ABB RAPID module: CalibData.mod

MODULE CalibData
    PERS tooldata My_Mechanism_1:=[TRUE,[[0,0,90],[1,0,0,0]],[1,[0,0,90],[1,0,0,0],0,0,0]];
    TASK PERS wobjdata Workobject_2:=[FALSE,TRUE,"",[[0,0,0],[1,0,0,0]],[[0,0,0],[1,0,0,0]]];
    TASK PERS wobjdata Workobject_3:=[FALSE,TRUE,"",[[1970.926,882.727,800],[1,0,0,0]],[[0,0,0],[1,0,0,0]]];
ENDMODULE
